(* IEC 61131-3 sources: codesys-framework/txt/application/WeVe Core (library)/60 Event/FB_Event/Properties, 5 files *)

(* ---- Active.prop.st ---- *)
PROPERTY Active : BOOL
// --- BEGIN IMPLEMENTATION ---

// ----------- GET -----------
VAR
END_VAR

// -- BEGIN IMPLEMENTATION GET --
Active := _xActive;

(* ---- Config.prop.st ---- *)
PROPERTY Config : SC_Event
// --- BEGIN IMPLEMENTATION ---

// ----------- GET -----------
VAR
END_VAR

// -- BEGIN IMPLEMENTATION GET --
Config := _scConfig;

// ----------- SET -----------
PUBLIC
VAR
END_VAR

// -- BEGIN IMPLEMENTATION SET --
_scConfig := Config;

(* ---- Disabled.prop.st ---- *)
PROPERTY Disabled : BOOL
// --- BEGIN IMPLEMENTATION ---

// ----------- GET -----------
VAR
END_VAR

// -- BEGIN IMPLEMENTATION GET --
Disabled := _xDisabled;

// ----------- SET -----------
PUBLIC
VAR
END_VAR

// -- BEGIN IMPLEMENTATION SET --
_xDisabled := Disabled;

// Uitgeschakeld event is nooit actief
IF _xDisabled THEN
	_xActive := FALSE;
	_xCondition := FALSE;
END_IF

(* ---- Level.prop.st ---- *)
PROPERTY Level : E_EventLevels
// --- BEGIN IMPLEMENTATION ---

// ----------- GET -----------
VAR
END_VAR

// -- BEGIN IMPLEMENTATION GET --
Level := _scConfig.eEventLevel;

(* ---- Logger.prop.st ---- *)
PROPERTY Logger : I_Logger
// --- BEGIN IMPLEMENTATION ---

// ----------- SET -----------
PUBLIC
VAR
END_VAR

// -- BEGIN IMPLEMENTATION SET --
_fbLogger := Logger;
